(* IEC 61131-3 sources: plc-iiot-stack/src/POUs/Iiot/FB_MqttTelemetry, 12 files *)

(* ---- FB_MqttTelemetry.decl.st ---- *)
// Назначение: публикация телеметрии (data_schema 3): одна метрика — один топик <prefix>/<device>/<metric>,
//             JSON {schema_version, ts, value, quality, unit}, QoS 1, retain. По изменению: Analog — когда
//             значение ушло от опубликованного больше зоны нечувствительности, Integer — при любом изменении
//             (зона 0), не чаще tMinInterval на метрику; смена quality — сразу. Контрольная публикация всех
//             метрик — раз в tPeriod и после каждого рождения узла (xReady). За вызов — не больше
//             uiMaxPerCycle публикаций, обход по кругу: ни одна метрика не ждёт вечно.
// Автор:      kr0nsch
// Версия:     0.1.1
// Документ:   docs/plc_mqtt.md, раздел «Телеметрия»
FUNCTION_BLOCK FB_MqttTelemetry
VAR_INPUT
    xEnable : BOOL;
    xReady : BOOL;                                           // связь есть и рождение опубликовано (FB_MqttDiag)
    itfClient : I_MqttClient;
    ltNow : LTIME;                                           // монотонное время (LTIME())
    uliTs_ms : ULINT;                                        // время UTC, мс от 1970 (поле ts)
    sTopicPrefix : STRING(GVL_Const.IIOT_PREFIX_LEN);        // site/area/unit
    tPeriod : TIME := GVL_Const.TELEMETRY_PERIOD_DEFAULT;   // T#0S — без контрольной публикации
    tMinInterval : TIME := GVL_Const.TELEMETRY_MIN_INTERVAL;
    uiMaxPerCycle : UINT := GVL_Const.TELEMETRY_MAX_PER_CYCLE;
END_VAR
VAR_IN_OUT
    aPoints : ARRAY[*] OF ST_IiotPoint;
END_VAR
VAR_OUTPUT
    udiPublished : UDINT;       // принято клиентом
    udiFailed : UDINT;          // клиент не принял (нет места в очереди): метрика повторится
    udiDropped : UDINT;         // JSON или топик не поместились: метрика пропущена
    uiPending : UINT;           // метрик ждут публикации после этого вызова
END_VAR
VAR
    fbJson : FB_JsonBuilder;
    sTopic : STRING(GVL_Const.MQTT_TOPIC_LEN);
    xPeriodRunning : BOOL;
    ltPeriodStart : LTIME;
    diCursor : DINT;            // с какой метрики начинать обход в следующем вызове
END_VAR

(* ---- FB_MqttTelemetry.impl.st ---- *)
// Нет связи или рождения: после него всё публикуется заново
IF NOT xEnable OR NOT xReady OR itfClient = 0 OR NOT F_IiotClockValid(uliTs_ms := uliTs_ms) THEN
    ResetSent(aPointTable := aPoints);
    RETURN;
END_IF
IF NOT itfClient.IsConnected() THEN
    ResetSent(aPointTable := aPoints);
    RETURN;
END_IF

// Контрольная публикация: все метрики принудительно
IF NOT xPeriodRunning OR ltNow < ltPeriodStart THEN
    xPeriodRunning := TRUE;
    ltPeriodStart := ltNow;
ELSIF tPeriod > T#0S AND_THEN (ltNow - ltPeriodStart) >= TIME_TO_LTIME(tPeriod) THEN
    ltPeriodStart := ltNow;
    ForceAll(aPointTable := aPoints);
END_IF

PublishDue(aPointTable := aPoints);

(* ---- ForceAll.method.decl.st ---- *)
// Пометить все метрики для контрольной публикации.
METHOD PRIVATE ForceAll
VAR_IN_OUT
    aPointTable : ARRAY[*] OF ST_IiotPoint;
END_VAR
VAR
    diIdx : DINT;
END_VAR

(* ---- ForceAll.method.impl.st ---- *)
FOR diIdx := LOWER_BOUND(aPointTable, 1) TO UPPER_BOUND(aPointTable, 1) DO
    aPointTable[diIdx].xForce := TRUE;
END_FOR

(* ---- PointDue.method.decl.st ---- *)
// Нужна ли публикация: не публиковалась с подключения, контрольная, сменилось качество — сразу; изменение
// значения — не раньше tMinInterval после прошлой публикации (метрики xPeriodicOnly — только контрольно).
METHOD PRIVATE PointDue : BOOL
VAR_IN_OUT CONSTANT
    // lint:allow STL007 параметр VAR_IN_OUT CONSTANT — ссылка только для чтения, а не константа
    stPoint : ST_IiotPoint;
END_VAR

(* ---- PointDue.method.impl.st ---- *)
IF NOT stPoint.xSent OR stPoint.xForce OR stPoint.eQuality <> stPoint.eLastQuality THEN
    PointDue := TRUE;
    RETURN;
END_IF
IF stPoint.stCfg.xPeriodicOnly THEN
    RETURN;
END_IF
IF ltNow >= stPoint.ltLastSent AND_THEN (ltNow - stPoint.ltLastSent) < TIME_TO_LTIME(tMinInterval) THEN
    RETURN;
END_IF
PointDue := F_IiotDeadbandExceeded(lrNew := stPoint.lrValue, lrLast := stPoint.lrLastValue,
                                   rDeadband := stPoint.stCfg.rDeadband);

(* ---- PublishDue.method.decl.st ---- *)
// Обход метрик по кругу от diCursor: опубликовать те, что требуют публикации, не больше uiMaxPerCycle.
// Клиент отказал — публикации до следующего вызова прекращаются. uiPending — сколько метрик ждут.
METHOD PRIVATE PublishDue
VAR_IN_OUT
    aPointTable : ARRAY[*] OF ST_IiotPoint;
END_VAR
VAR
    diLo : DINT;
    diTotal : DINT;
    diStep : DINT;
    diIdx : DINT;
    diNextCursor : DINT;
    uiBudget : UINT;
    xBlocked : BOOL;        // клиент не принял сообщение в этом вызове
END_VAR

(* ---- PublishDue.method.impl.st ---- *)
diLo := LOWER_BOUND(aPointTable, 1);
diTotal := UPPER_BOUND(aPointTable, 1) - diLo + 1;
uiPending := 0;
IF diTotal <= 0 THEN
    RETURN;
END_IF
IF diCursor < 0 OR diCursor >= diTotal THEN
    diCursor := 0;
END_IF
uiBudget := MAX(uiMaxPerCycle, 1);
diNextCursor := -1;
FOR diStep := 0 TO diTotal - 1 DO
    diIdx := diLo + (diCursor + diStep) MOD diTotal;
    IF PointDue(stPoint := aPointTable[diIdx]) THEN
        IF uiBudget > 0 AND NOT xBlocked THEN
            IF PublishPoint(stPoint := aPointTable[diIdx]) THEN
                uiBudget := uiBudget - 1;
            ELSE
                xBlocked := TRUE;
            END_IF
        END_IF
        IF PointDue(stPoint := aPointTable[diIdx]) THEN
            uiPending := uiPending + 1;
            IF diNextCursor < 0 THEN
                diNextCursor := diIdx - diLo;   // здесь начнём в следующем вызове
            END_IF
        END_IF
    END_IF
END_FOR
IF diNextCursor >= 0 THEN
    diCursor := diNextCursor;
END_IF

(* ---- PublishPoint.method.decl.st ---- *)
// Опубликовать метрику: {"schema_version","ts","value","quality"[,"unit"]}. TRUE — метрика обработана
// (опубликована или пропущена из-за переполнения); FALSE — клиент не принял, она повторится.
// Значение не конечно (NaN, ±Inf): схема требует число, поэтому передаётся последнее опубликованное
// конечное значение с quality = bad (data_schema 3.2).
METHOD PRIVATE PublishPoint : BOOL
VAR_IN_OUT
    stPoint : ST_IiotPoint;
END_VAR
VAR
    xFinite : BOOL;
    lrOut : LREAL;
    eOutQuality : E_IiotQuality;
END_VAR

(* ---- PublishPoint.method.impl.st ---- *)
sTopic := F_IiotTopic(sPrefix := sTopicPrefix, sPath := stPoint.stCfg.sPath);
xFinite := F_IsFiniteLreal(lrValue := stPoint.lrValue);
IF xFinite THEN
    lrOut := stPoint.lrValue;
    eOutQuality := stPoint.eQuality;
ELSE
    lrOut := stPoint.lrLastFinite;
    eOutQuality := E_IiotQuality.Bad;
END_IF
fbJson.Begin();
fbJson.AddString(sKey := 'schema_version', sValue := GVL_Const.IIOT_SCHEMA_VERSION);
fbJson.AddInt(sKey := 'ts', liValue := ULINT_TO_LINT(uliTs_ms));
IF stPoint.stCfg.eKind = E_IiotValueKind.Analog THEN
    fbJson.AddReal(sKey := 'value', lrValue := lrOut, uiDecimals := stPoint.stCfg.uiDecimals);
ELSE
    fbJson.AddInt(sKey := 'value', liValue := LREAL_TO_LINT(lrOut));
END_IF
fbJson.AddString(sKey := 'quality', sValue := F_IiotQualityText(eQuality := eOutQuality));
IF LEN(stPoint.stCfg.sUnit) > 0 THEN
    fbJson.AddString(sKey := 'unit', sValue := stPoint.stCfg.sUnit);
END_IF

IF NOT fbJson.Finish() OR LEN(sTopic) = 0 THEN
    udiDropped := udiDropped + 1;     // повторять бессмысленно: размер не изменится
ELSIF itfClient.Publish(sTopic := sTopic, eQos := E_MqttQos.AtLeastOnce, xRetain := TRUE,
                        sPayload := fbJson.sJson) THEN
    udiPublished := udiPublished + 1;
ELSE
    udiFailed := udiFailed + 1;
    RETURN;
END_IF
stPoint.lrLastValue := stPoint.lrValue;
IF xFinite THEN
    stPoint.lrLastFinite := stPoint.lrValue;
END_IF
stPoint.eLastQuality := stPoint.eQuality;
stPoint.ltLastSent := ltNow;
stPoint.xSent := TRUE;
stPoint.xForce := FALSE;
PublishPoint := TRUE;

(* ---- ResetSent.method.decl.st ---- *)
// Связи нет: сбросить признаки «опубликовано», чтобы после рождения опубликовать всё; период — заново.
METHOD PRIVATE ResetSent
VAR_IN_OUT
    aPointTable : ARRAY[*] OF ST_IiotPoint;
END_VAR
VAR
    diIdx : DINT;
END_VAR

(* ---- ResetSent.method.impl.st ---- *)
FOR diIdx := LOWER_BOUND(aPointTable, 1) TO UPPER_BOUND(aPointTable, 1) DO
    aPointTable[diIdx].xSent := FALSE;
END_FOR
xPeriodRunning := FALSE;
uiPending := 0;
